// TIA Portal V21 export
// export: Created 2026-11-10T07:35:22.8631173Z, ExportSetting WithDefaults, DisplayName Totally Integrated Automation Portal, DisplayVersion V21 Update 3, DisplayName STEP 7 Professional, DisplayVersion V21 Update 3, DisplayName STEP 7 Safety, DisplayVersion V21, DisplayName Tech WebApplication, DisplayVersion V21, DisplayName WinCC Basic/Comfort/Advanced, DisplayVersion V21 Update 3, DisplayName WinCC Unified, DisplayVersion V21 Update 3
FUNCTION_BLOCK "FB_Lad_ex153"   // FB193, LAD
{ S7_Optimized_Access := 'TRUE' }
VERSION : 0.1
// stored: AutoNumber true, IsIECCheckEnabled false, IsRetainMemResEnabled false, MemoryReserve 100, SetENOAutomatically false, UDAEnableTagReadback false
   VAR_INPUT
      v_laddr : HW_ANY;
   END_VAR
   VAR_OUTPUT
      v_ret_val : Int;
   END_VAR
   VAR_IN_OUT
      v_geoaddr : GEOADDR;
   END_VAR
BEGIN

REGION Network 1: LOG2GEO - Determine slot from hardware identifier
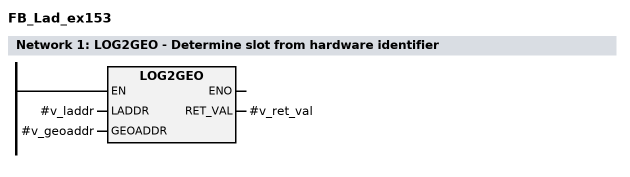
   RUNG wire#powerrail
      LOG2GEO(LADDR := #v_laddr, Ret_Val => #v_ret_val, GEOADDR := #v_geoaddr)
   END_RUNG
   // the same network as SCL:
   #v_ret_val := LOG2GEO(LADDR := #v_laddr, GEOADDR := #v_geoaddr);
END_REGION
END_FUNCTION_BLOCK
